// TIA Portal project "2026_10_13_Imbottigliatrice" (V15)

(* hardware
DEVICE "S7-1200 station_1"  S7-1200 Station
   slot 0: "Telaio di montaggio_0"  S7-1200 Rack  Rack  V1.0
   slot 1: "PLC_1"  CPU 1215C DC/DC/DC  6ES7 215-1AG40-0XB0  V4.2
*)

// ===== PLC "PLC_1"  CPU 1215C DC/DC/DC =====

VAR_GLOBAL   // PLC tag table "Tabella delle variabili standard"
   "System_Byte" AT %MB1 : Byte;
   "FirstScan" AT %M1.0 : Bool;
   "DiagStatusUpdate" AT %M1.1 : Bool;
   "AlwaysTRUE" AT %M1.2 : Bool;
   "AlwaysFALSE" AT %M1.3 : Bool;
   "Clock_Byte" AT %MB0 : Byte;
   "Clock_10Hz" AT %M0.0 : Bool;
   "Clock_5Hz" AT %M0.1 : Bool;
   "Clock_2.5Hz" AT %M0.2 : Bool;
   "Clock_2Hz" AT %M0.3 : Bool;
   "Clock_1.25Hz" AT %M0.4 : Bool;
   "Clock_1Hz" AT %M0.5 : Bool;
   "Clock_0.625Hz" AT %M0.6 : Bool;
   "Clock_0.5Hz" AT %M0.7 : Bool;
END_VAR

VAR_GLOBAL   // PLC tag table "Ingressi"
   "IC" AT %I0.0 : Bool;   // Pulsante di inizio ciclo
   "FC" AT %I0.1 : Bool;   // Pulsante di STOP/Emergenza (NC)
   "Fc0" AT %I0.2 : Bool;   // Sensore di prossimità (pos iniziale)
   "Fc1" AT %I0.3 : Bool;   // Sensore di prossimità (pos riempimento)
   "Fc2" AT %I0.4 : Bool;   // Sensore di prossimità (pos tappatura)
   "Fc3" AT %I0.5 : Bool;   // Sensore di prossimità (pos finale)
   "Fcs" AT %I0.6 : Bool;   // Sensore di prossimità (presenza scatola)
   "SL" AT %I0.7 : Bool;   // Sensore di prossimità (livello composto)
   "a0" AT %I1.0 : Bool;   // Fine corsa cilindro A chiuso
   "a1" AT %I1.1 : Bool;   // Fine corsa cilindro A aperto
   "b0" AT %I1.2 : Bool;   // Fine corsa cilindro B chiuso
   "b1" AT %I1.3 : Bool;   // Fine corsa cilindro B aperto
   "c0" AT %I1.4 : Bool;   // Fine corsa cilindro C chiuso
   "c1" AT %I1.5 : Bool;   // Fine corsa cilindro C aperto
END_VAR

VAR_GLOBAL   // PLC tag table "Uscite"
   "KM1" AT %Q0.0 : Bool;   // Teleruttore attivazione motore M1
   "Kev" AT %Q0.1 : Bool;   // Elettrovalvola erogazione composto
   "A+" AT %Q0.2 : Bool;   // Corsa positiva cilindro A (bistabile)
   "A-" AT %Q0.3 : Bool;   // Corsa negativa cilndro A (bistabile)
   "B+" AT %Q0.4 : Bool;   // Corsa positiva cilindro B (bistabile)
   "B-" AT %Q0.5 : Bool;   // Corsa negatica cilindro B (bistabile)
   "C+" AT %Q0.6 : Bool;   // Corsa positiva cilindro C (monostabile)
   "HLL" AT %Q0.7 : Bool;   // Segnalazione lampeggiante impianto in funzionamento
   "HLPi" AT %Q1.0 : Bool;   // Presenza bottiglia inizio nastro
   "HLPf" AT %Q1.1 : Bool;   // Presenza bottiglia fine nastro
   "HLM1" AT %M20.0 : Bool;   // Segnalazione motore M1 (virtuale)
   "HLE" AT %M20.1 : Bool;   // Segnalazione estrusione (virtuale)
   "HLB" AT %M20.2 : Bool;   // Segnalazione blocco bottiglia (virtuale)
   "HLC" AT %M20.3 : Bool;   // Segnalazione tappatura (virtuale)
   "HLSF" AT %M20.4 : Bool;   // Segnalazione scatola piena (virtuale)
END_VAR

VAR_GLOBAL   // PLC tag table "Merker"
   "FASE" AT %MW100 : Int;   // Variabile di stato
   "n" AT %MW102 : Int;   // Variabile di conteggio
END_VAR

// folder: System blocks/Program resources

DATA_BLOCK "TON_0"   // DB1
{ S7_Optimized_Access := 'TRUE' }
AUTHOR : Simatic
FAMILY : IEC
NAME : IEC_TMR
VERSION : 1.0
// stored: InstanceOfName IEC_TIMER
"IEC_TIMER"
BEGIN
END_DATA_BLOCK

DATA_BLOCK "CTU_0"   // DB2
{ S7_Optimized_Access := 'TRUE' }
AUTHOR : Simatic
FAMILY : IEC
NAME : CNTR
VERSION : 1.0
// stored: InstanceOfName IEC_COUNTER
"IEC_COUNTER"
BEGIN
END_DATA_BLOCK

// folder: (top level)

FUNCTION "Controllo" : Void   // FC1, LAD
{ S7_Optimized_Access := 'TRUE' }
VERSION : 0.1
   VAR_TEMP   // added for the SCL form of the ladder/FBD networks
      _w1 : Bool;
   END_VAR
BEGIN

REGION Network 1: Attesa inizio ciclo
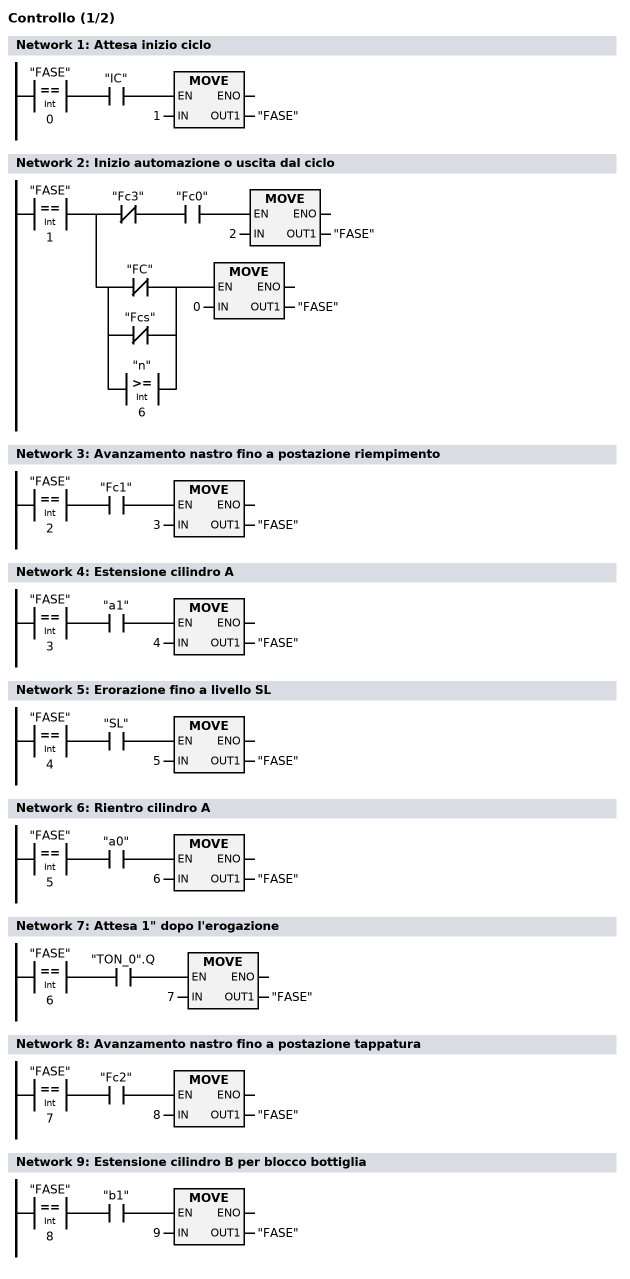
   RUNG wire#powerrail
      { S7_Templates := "SrcType := Int" } EQ_Contact(in1 := "FASE", in2 := 0)
      Contact( "IC" )
      Move(in := 1, out1 => "FASE")
   END_RUNG
   // the same network as SCL:
   IF ("FASE" = 0) AND "IC" THEN "FASE" := 1; END_IF;
END_REGION

REGION Network 2: Inizio automazione o uscita dal ciclo
   RUNG wire#powerrail
      { S7_Templates := "SrcType := Int" } EQ_Contact(in1 := "FASE", in2 := 1)
      wire#w1
      I_Contact( "Fc3" )
      Contact( "Fc0" )
      Move(in := 2, out1 => "FASE")
   END_RUNG
   RUNG wire#w1
      I_Contact( "FC" )
      wire#w2
      Move(in := 0, out1 => "FASE")
   END_RUNG
   RUNG wire#w1
      I_Contact( "Fcs" )
   END_RUNG wire#w2
   RUNG wire#w1
      { S7_Templates := "SrcType := Int" } GE_Contact(in1 := "n", in2 := 6)
   END_RUNG wire#w2
   // the same network as SCL:
   #_w1 := "FASE" = 1;
   IF #_w1 AND NOT "Fc3" AND "Fc0" THEN "FASE" := 2; END_IF;
   IF #_w1 AND (NOT "FC" OR NOT "Fcs" OR ("n" >= 6)) THEN "FASE" := 0; END_IF;
END_REGION

REGION Network 3: Avanzamento nastro fino a postazione riempimento
   RUNG wire#powerrail
      { S7_Templates := "SrcType := Int" } EQ_Contact(in1 := "FASE", in2 := 2)
      Contact( "Fc1" )
      Move(in := 3, out1 => "FASE")
   END_RUNG
   // the same network as SCL:
   IF ("FASE" = 2) AND "Fc1" THEN "FASE" := 3; END_IF;
END_REGION

REGION Network 4: Estensione cilindro A
   RUNG wire#powerrail
      { S7_Templates := "SrcType := Int" } EQ_Contact(in1 := "FASE", in2 := 3)
      Contact( "a1" )
      Move(in := 4, out1 => "FASE")
   END_RUNG
   // the same network as SCL:
   IF ("FASE" = 3) AND "a1" THEN "FASE" := 4; END_IF;
END_REGION

REGION Network 5: Erorazione fino a livello SL
   RUNG wire#powerrail
      { S7_Templates := "SrcType := Int" } EQ_Contact(in1 := "FASE", in2 := 4)
      Contact( "SL" )
      Move(in := 5, out1 => "FASE")
   END_RUNG
   // the same network as SCL:
   IF ("FASE" = 4) AND "SL" THEN "FASE" := 5; END_IF;
END_REGION

REGION Network 6: Rientro cilindro A
   RUNG wire#powerrail
      { S7_Templates := "SrcType := Int" } EQ_Contact(in1 := "FASE", in2 := 5)
      Contact( "a0" )
      Move(in := 6, out1 => "FASE")
   END_RUNG
   // the same network as SCL:
   IF ("FASE" = 5) AND "a0" THEN "FASE" := 6; END_IF;
END_REGION

REGION Network 7: Attesa 1" dopo l'erogazione
   RUNG wire#powerrail
      { S7_Templates := "SrcType := Int" } EQ_Contact(in1 := "FASE", in2 := 6)
      Contact( "TON_0".Q )
      Move(in := 7, out1 => "FASE")
   END_RUNG
   // the same network as SCL:
   IF ("FASE" = 6) AND "TON_0".Q THEN "FASE" := 7; END_IF;
END_REGION

REGION Network 8: Avanzamento nastro fino a postazione tappatura
   RUNG wire#powerrail
      { S7_Templates := "SrcType := Int" } EQ_Contact(in1 := "FASE", in2 := 7)
      Contact( "Fc2" )
      Move(in := 8, out1 => "FASE")
   END_RUNG
   // the same network as SCL:
   IF ("FASE" = 7) AND "Fc2" THEN "FASE" := 8; END_IF;
END_REGION

REGION Network 9: Estensione cilindro B per blocco bottiglia
   RUNG wire#powerrail
      { S7_Templates := "SrcType := Int" } EQ_Contact(in1 := "FASE", in2 := 8)
      Contact( "b1" )
      Move(in := 9, out1 => "FASE")
   END_RUNG
   // the same network as SCL:
   IF ("FASE" = 8) AND "b1" THEN "FASE" := 9; END_IF;
END_REGION

REGION Network 10: Estensione cilindro C per tappatura
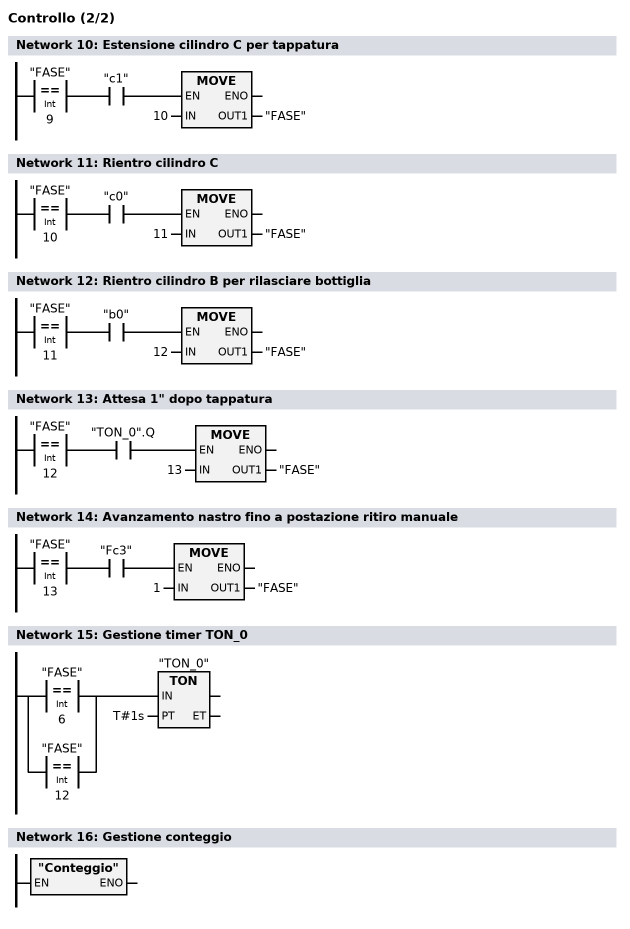
   RUNG wire#powerrail
      { S7_Templates := "SrcType := Int" } EQ_Contact(in1 := "FASE", in2 := 9)
      Contact( "c1" )
      Move(in := 10, out1 => "FASE")
   END_RUNG
   // the same network as SCL:
   IF ("FASE" = 9) AND "c1" THEN "FASE" := 10; END_IF;
END_REGION

REGION Network 11: Rientro cilindro C
   RUNG wire#powerrail
      { S7_Templates := "SrcType := Int" } EQ_Contact(in1 := "FASE", in2 := 10)
      Contact( "c0" )
      Move(in := 11, out1 => "FASE")
   END_RUNG
   // the same network as SCL:
   IF ("FASE" = 10) AND "c0" THEN "FASE" := 11; END_IF;
END_REGION

REGION Network 12: Rientro cilindro B per rilasciare bottiglia
   RUNG wire#powerrail
      { S7_Templates := "SrcType := Int" } EQ_Contact(in1 := "FASE", in2 := 11)
      Contact( "b0" )
      Move(in := 12, out1 => "FASE")
   END_RUNG
   // the same network as SCL:
   IF ("FASE" = 11) AND "b0" THEN "FASE" := 12; END_IF;
END_REGION

REGION Network 13: Attesa 1" dopo tappatura
   RUNG wire#powerrail
      { S7_Templates := "SrcType := Int" } EQ_Contact(in1 := "FASE", in2 := 12)
      Contact( "TON_0".Q )
      Move(in := 13, out1 => "FASE")
   END_RUNG
   // the same network as SCL:
   IF ("FASE" = 12) AND "TON_0".Q THEN "FASE" := 13; END_IF;
END_REGION

REGION Network 14: Avanzamento nastro fino a postazione ritiro manuale
   RUNG wire#powerrail
      { S7_Templates := "SrcType := Int" } EQ_Contact(in1 := "FASE", in2 := 13)
      Contact( "Fc3" )
      Move(in := 1, out1 => "FASE")
   END_RUNG
   // the same network as SCL:
   IF ("FASE" = 13) AND "Fc3" THEN "FASE" := 1; END_IF;
END_REGION

REGION Network 15: Gestione timer TON_0
   "TON_0".TON(IN := ("FASE" = 6) OR ("FASE" = 12), PT := T#1s);
END_REGION

REGION Network 16: Gestione conteggio
   RUNG wire#powerrail
      "Conteggio"()
   END_RUNG
   // the same network as SCL:
   "Conteggio"();
END_REGION
END_FUNCTION

FUNCTION "Comando" : Void   // FC2, LAD
{ S7_Optimized_Access := 'TRUE' }
VERSION : 0.1
BEGIN

REGION Network 1: Azionamento motore M1
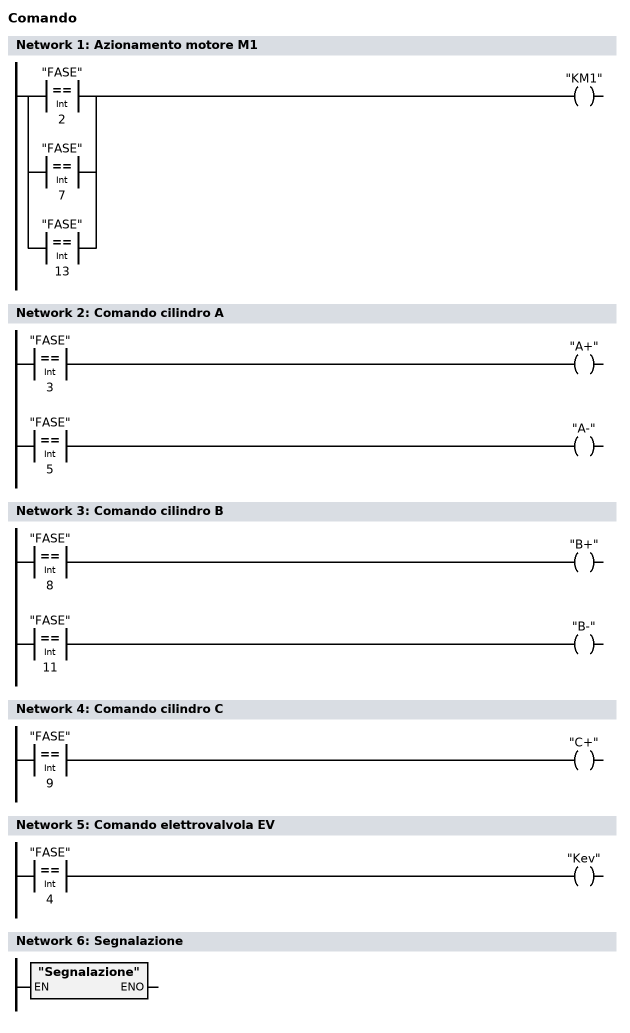
   RUNG wire#powerrail
      { S7_Templates := "SrcType := Int" } EQ_Contact(in1 := "FASE", in2 := 2)
      wire#w1
      Coil( "KM1" )
   END_RUNG
   RUNG wire#powerrail
      { S7_Templates := "SrcType := Int" } EQ_Contact(in1 := "FASE", in2 := 7)
   END_RUNG wire#w1
   RUNG wire#powerrail
      { S7_Templates := "SrcType := Int" } EQ_Contact(in1 := "FASE", in2 := 13)
   END_RUNG wire#w1
   // the same network as SCL:
   "KM1" := ("FASE" = 2) OR ("FASE" = 7) OR ("FASE" = 13);
END_REGION

REGION Network 2: Comando cilindro A
   RUNG wire#powerrail
      { S7_Templates := "SrcType := Int" } EQ_Contact(in1 := "FASE", in2 := 3)
      Coil( "A+" )
   END_RUNG
   RUNG wire#powerrail
      { S7_Templates := "SrcType := Int" } EQ_Contact(in1 := "FASE", in2 := 5)
      Coil( "A-" )
   END_RUNG
   // the same network as SCL:
   "A+" := "FASE" = 3;
   "A-" := "FASE" = 5;
END_REGION

REGION Network 3: Comando cilindro B
   RUNG wire#powerrail
      { S7_Templates := "SrcType := Int" } EQ_Contact(in1 := "FASE", in2 := 8)
      Coil( "B+" )
   END_RUNG
   RUNG wire#powerrail
      { S7_Templates := "SrcType := Int" } EQ_Contact(in1 := "FASE", in2 := 11)
      Coil( "B-" )
   END_RUNG
   // the same network as SCL:
   "B+" := "FASE" = 8;
   "B-" := "FASE" = 11;
END_REGION

REGION Network 4: Comando cilindro C
   RUNG wire#powerrail
      { S7_Templates := "SrcType := Int" } EQ_Contact(in1 := "FASE", in2 := 9)
      Coil( "C+" )
   END_RUNG
   // the same network as SCL:
   "C+" := "FASE" = 9;
END_REGION

REGION Network 5: Comando elettrovalvola EV
   RUNG wire#powerrail
      { S7_Templates := "SrcType := Int" } EQ_Contact(in1 := "FASE", in2 := 4)
      Coil( "Kev" )
   END_RUNG
   // the same network as SCL:
   "Kev" := "FASE" = 4;
END_REGION

REGION Network 6: Segnalazione
   RUNG wire#powerrail
      "Segnalazione"()
   END_RUNG
   // the same network as SCL:
   "Segnalazione"();
END_REGION
END_FUNCTION

FUNCTION "Conteggio" : Void   // FC4, LAD
{ S7_Optimized_Access := 'TRUE' }
VERSION : 0.1
BEGIN

REGION Network 1: Incremento conteggio con rimozione bottiglia, Reset con rimozione scatola
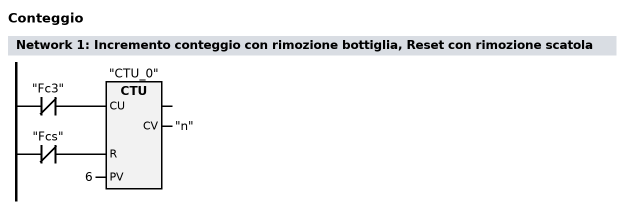
   "CTU_0".CTU(CU := NOT "Fc3", R := NOT "Fcs", PV := 6, CV => "n");
END_REGION
END_FUNCTION

FUNCTION "Segnalazione" : Void   // FC5, LAD
{ S7_Optimized_Access := 'TRUE' }
VERSION : 0.1
BEGIN

REGION Network 1: Lampeggio
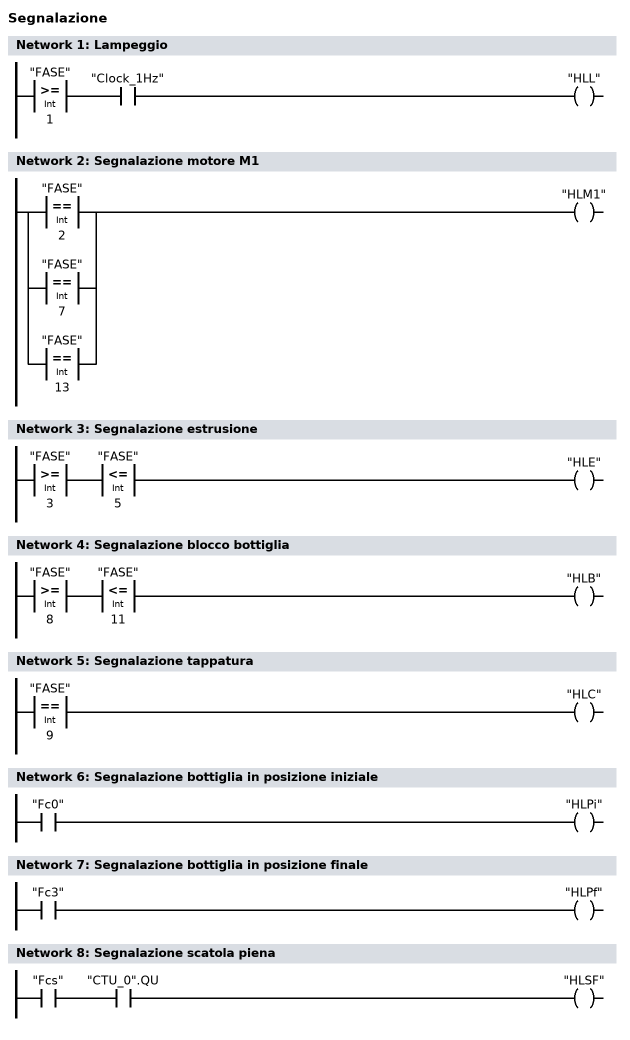
   RUNG wire#powerrail
      { S7_Templates := "SrcType := Int" } GE_Contact(in1 := "FASE", in2 := 1)
      Contact( "Clock_1Hz" )
      Coil( "HLL" )
   END_RUNG
   // the same network as SCL:
   "HLL" := ("FASE" >= 1) AND "Clock_1Hz";
END_REGION

REGION Network 2: Segnalazione motore M1
   RUNG wire#powerrail
      { S7_Templates := "SrcType := Int" } EQ_Contact(in1 := "FASE", in2 := 2)
      wire#w1
      Coil( "HLM1" )
   END_RUNG
   RUNG wire#powerrail
      { S7_Templates := "SrcType := Int" } EQ_Contact(in1 := "FASE", in2 := 7)
   END_RUNG wire#w1
   RUNG wire#powerrail
      { S7_Templates := "SrcType := Int" } EQ_Contact(in1 := "FASE", in2 := 13)
   END_RUNG wire#w1
   // the same network as SCL:
   "HLM1" := ("FASE" = 2) OR ("FASE" = 7) OR ("FASE" = 13);
END_REGION

REGION Network 3: Segnalazione estrusione
   RUNG wire#powerrail
      { S7_Templates := "SrcType := Int" } GE_Contact(in1 := "FASE", in2 := 3)
      { S7_Templates := "SrcType := Int" } LE_Contact(in1 := "FASE", in2 := 5)
      Coil( "HLE" )
   END_RUNG
   // the same network as SCL:
   "HLE" := ("FASE" >= 3) AND ("FASE" <= 5);
END_REGION

REGION Network 4: Segnalazione blocco bottiglia
   RUNG wire#powerrail
      { S7_Templates := "SrcType := Int" } GE_Contact(in1 := "FASE", in2 := 8)
      { S7_Templates := "SrcType := Int" } LE_Contact(in1 := "FASE", in2 := 11)
      Coil( "HLB" )
   END_RUNG
   // the same network as SCL:
   "HLB" := ("FASE" >= 8) AND ("FASE" <= 11);
END_REGION

REGION Network 5: Segnalazione tappatura
   RUNG wire#powerrail
      { S7_Templates := "SrcType := Int" } EQ_Contact(in1 := "FASE", in2 := 9)
      Coil( "HLC" )
   END_RUNG
   // the same network as SCL:
   "HLC" := "FASE" = 9;
END_REGION

REGION Network 6: Segnalazione bottiglia in posizione iniziale
   RUNG wire#powerrail
      Contact( "Fc0" )
      Coil( "HLPi" )
   END_RUNG
   // the same network as SCL:
   "HLPi" := "Fc0";
END_REGION

REGION Network 7: Segnalazione bottiglia in posizione finale
   RUNG wire#powerrail
      Contact( "Fc3" )
      Coil( "HLPf" )
   END_RUNG
   // the same network as SCL:
   "HLPf" := "Fc3";
END_REGION

REGION Network 8: Segnalazione scatola piena
   RUNG wire#powerrail
      Contact( "Fcs" )
      Contact( "CTU_0".QU )
      Coil( "HLSF" )
   END_RUNG
   // the same network as SCL:
   "HLSF" := "Fcs" AND "CTU_0".QU;
END_REGION
END_FUNCTION

ORGANIZATION_BLOCK "Main"   // OB1, LAD, ProgramCycle
TITLE = "Main Program Sweep (Cycle)"
{ S7_Optimized_Access := 'TRUE' }
VERSION : 0.1
   VAR_INPUT
      Initial_Call : Bool;   // Initial call of this OB
      Remanence : Bool;   // =True, if remanent data are available
   END_VAR
BEGIN

REGION Network 1: Controllo
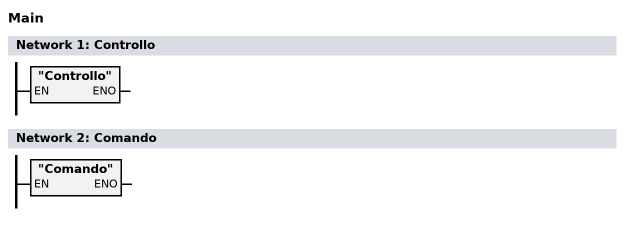
   RUNG wire#powerrail
      "Controllo"()
   END_RUNG
   // the same network as SCL:
   "Controllo"();
END_REGION

REGION Network 2: Comando
   RUNG wire#powerrail
      "Comando"()
   END_RUNG
   // the same network as SCL:
   "Comando"();
END_REGION
END_ORGANIZATION_BLOCK

ORGANIZATION_BLOCK "Startup"   // OB100, LAD, Startup
TITLE = "Complete Restart"
{ S7_Optimized_Access := 'TRUE' }
VERSION : 0.1
   VAR_INPUT
      LostRetentive : Bool;   // True if retentive data are lost
      LostRTC : Bool;   // True if date and time are lost
   END_VAR
BEGIN

REGION Network 1: Reset stato iniziale
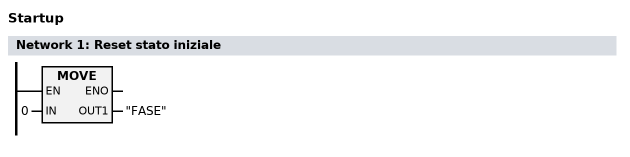
   RUNG wire#powerrail
      Move(in := 0, out1 => "FASE")
   END_RUNG
   // the same network as SCL:
   "FASE" := 0;
END_REGION
END_ORGANIZATION_BLOCK